Staubli VAL3: HMI_pointEdit.pjx

--- HMI_pointEdit.pjx ---
Parameters version=s8.15.3Cs9_BS3337 stackSize=5000 millimeterUnit=true
Program file=bind.pgx
Program file=insertAction.pgx
Program file=insertDelay.pgx
Program file=insertDelay1.pgx
Program file=insertIF.pgx
Program file=insertSignal.pgx
Program file=insertSwitch.pgx
Program file=load.pgx
Program file=main.pgx
Program file=onStart.pgx
Program file=paraBind.pgx
Program file=paraEdit.pgx
Program file=paraStart.pgx
Program file=refreshlist.pgx
Program file=sCommentIO.pgx
Program file=start.pgx
Program file=stop.pgx
Program file=teachPoint.pgx
Data file=HMI_pointEdit.dtx
Library alias=util path=Disk://HMI_cs9/HMI_util/HMI_util.pjx
Library alias=trajectory path=Disk://source/projectSource/trajectory/trajectory.pjx
Library alias=io path=Disk://source/projectSource/io/io.pjx
Library alias=savedata path=Disk://source/saveData/saveData.pjx
Library alias=actiondata path=Disk://data/actionData/actionData.pjx
Library alias=rs path=Disk://source/projectSource/robotStatus/robotStatus.pjx

--- HMI_pointEdit.dtx ---
mdesc mNomSpeed
bool bBack
string sTrajItem
string sUsingLib
string sUsingFrame
string sUsingTool
public bool bBool[30]
string sPageIndex
string sPageNum
public string sList = "0"
string sSelPoint
num nPageIndex
num nPageNum
bool bRefresh
bool bConfirm
bool bBackSignal
string sSignalType
string sSignalIndex
num nSignalValue
num nSignalType
string sLastType
string sIOList
bool bConfirmDelay
bool bBackDelay
num nSetDelay
public string sIFtype[3]
string sIFIndex[3]
public num nIOindex[3]
public num nIFvalue[3]
bool bConfirmIF
bool bBackIF
string sANDOR[2]
public num nANDOR[2]
num nIFtype[3]
num nParaSpeed
num nParaAccel
num nParaBlend
num nParaPercent
string sParaType
bool bParaJoint
bool bParaOFF
num nMoveType
bool bParaConfirm
bool bParaBack
bool bPAllModify
bool bLast
bool bToSave
frame fUsingFrame = {fatherId=world[0]}
tool tUsingTool = {fatherId=flange[0]}
public num nTRSF[12]
public string sTRSF[12]
string sBlendType
string sLastItem
string sLastMtype
num _nFrameID
num _nToolID
num _nPointIndex
string sComment
num nPointIndex
bool bSafePoint
string sActionList
bool bAConfirm
bool bACancel
string sSelAction
bool bConfirmSwitch
bool bBackSwitch
bool bMark
public string sCommentIO1
bool bToSave1
string sLastTrajItem
string sSelMovCPoint
bool bRecord
bool bMoveTo
bool bConfirmMovC
bool bCancelMovC
bool bShow2Point
string sParaPointType[2]

--- main.pgx ---
public program main(string x_sTrajItem)
  local bool l_bExit
  local num l_nPoint
  local bool l_bResult
  local num l_nPointSize
  local num l_nMoveType
  local bool l_bOperate
begin
  do
    if util:sPage!="point"
      util:sPage="point"
      call util:loadingPage()
      call onStart(x_sTrajItem)
      call trajectory:getFrameID(x_sTrajItem,_nFrameID)
      call trajectory:getToolID(x_sTrajItem,_nToolID)
      call refreshlist()
      call bind()
      userPage(util:sPage)
      delay(0.1)
      sLastItem=""
    endIf
    //point Move
    if workingMode()==1
      if sSelPoint!=sLastItem and sSelPoint!=""
        sLastItem=sSelPoint
        call trajectory:getPointIndex(sTrajItem,sSelPoint,l_nPoint,l_bResult)
        if !bMark
          if isPowered()
            //guohangxin modified 2023.03.23
            //            call trajectory:pointMove(sTrajItem,l_nPoint)
            if taskStatus("stepMove")>-1
              taskKill("stepMove")
              wait(taskStatus("stepMove")==-1)
            endIf
            taskCreate "stepMove",10,trajectory:pointMove(sTrajItem,l_nPoint)
          endIf
        else
          call trajectory:setMark(sTrajItem,l_nPoint)
          bRefresh=true
        endIf
      endIf
    endIf
    //button
    if bBool[0]
      //示教
      bBool[0]=false
      call trajectory:getPointIndex(sTrajItem,sSelPoint,l_nPoint,l_bResult)
      if l_bResult
        //call trajectory:teachPoint(sTrajItem,l_nPoint,bToSave)
        call teachPoint()
        bRefresh=true
      else
        userPageAlert("请选择有效点位！")
      endIf
    elseIf bBool[1]
      //标记
      bBool[1]=false
      bMark=!bMark
      if !bMark
        userPageSet("point","btn1","innerHTML","标记")
        call trajectory:resetMark(sTrajItem)
        bRefresh=true
      else
        userPageSet("point","btn1","innerHTML","取消标记")
        //call trajectory:resizeMark(sTrajItem)
      endIf
    elseIf bBool[2]
      bBool[2]=false
      //插入if
      call insertIF()
    elseIf bBool[3]
      bBool[3]=false
      //编辑
      call trajectory:getPointIndex(sTrajItem,sSelPoint,l_nPoint,l_bResult)
      if l_bResult
        call trajectory:getMoveType(sTrajItem,l_nPoint,l_nMoveType)
        if l_nMoveType==0 or l_nMoveType==1 or l_nMoveType==2
          call paraEdit()
        endIf
      else
        userPageAlert("未选择有效项！")
      endIf
    elseIf bBool[4]
      bBool[4]=false
      //插入点位
      call trajectory:getPointIndex(sTrajItem,sSelPoint,l_nPoint,l_bResult)
      if l_bResult
        call trajectory:insertPoint(sTrajItem,l_nPoint,bToSave)

      else
        call trajectory:getPointSize(sTrajItem,l_nPointSize)
        call trajectory:insertPoint(sTrajItem,l_nPointSize-1,bToSave)
      endIf
      bRefresh=true
    elseIf bBool[5]
      bBool[5]=false
      //删除
      call trajectory:getPointIndex(sTrajItem,sSelPoint,l_nPoint,l_bResult)
      if l_bResult
        call trajectory:deletePoint(sTrajItem,l_nPoint,bToSave)
      else
        userPageAlert("未选中有效点位")
      endIf
      bRefresh=true
    elseIf bBool[6]
      bBool[6]=false
      //插入信号
      call insertSignal()
      bRefresh=true
    elseIf bBool[7]
      bBool[7]=false
      //保存
      call trajectory:onSave(bToSave)
    elseIf bBool[8]
      bBool[8]=false
      //head page
      nPageIndex=0
      l_nPoint=0
      bRefresh=true
    elseIf bBool[9]
      //page up
      bBool[9]=false
      if nPageIndex>0
        nPageIndex=nPageIndex-1
        l_nPoint=0
      endIf
      bRefresh=true
    elseIf bBool[10]
      bBool[10]=false
      //page down
      if nPageIndex<nPageNum-1
        nPageIndex=nPageIndex+1
        l_nPoint=0
      endIf
      bRefresh=true
    elseIf bBool[11]
      //end page
      bBool[11]=false
      nPageIndex=nPageNum-1
      l_nPoint=0
      bRefresh=true
    elseIf bBool[12]
      bBool[12]=false
      call trajectory:getPointIndex(sTrajItem,sSelPoint,l_nPoint,l_bResult)
      if l_bResult
        call trajectory:insertENDIF(sTrajItem,l_nPoint,bToSave)
      else
        userPageAlert("未选中有效点位")
      endIf
      bRefresh=true
    elseIf bBool[13]
      bBool[13]=true
      //delay
      call insertDelay()
      bRefresh=true
    elseIf bBool[14]
      bBool[14]=false
      call trajectory:getPointIndex(sTrajItem,sSelPoint,l_nPoint,l_bResult)
      if l_bResult
        call trajectory:insertJoint(sTrajItem,l_nPoint,bToSave)
      else
        call trajectory:getPointSize(sTrajItem,l_nPointSize)
        call trajectory:insertJoint(sTrajItem,l_nPointSize-1,bToSave)
      endIf
      bRefresh=true
    elseIf bBool[15]
      bBool[15]=false
      call insertAction()
    elseIf bBool[16]
      //插入圆弧点位
      bBool[16]=false
      call trajectory:getPointIndex(sTrajItem,sSelPoint,l_nPoint,l_bResult)
      if l_bResult
        call trajectory:insertCirclePoint(sTrajItem,l_nPoint,bToSave)
      else
        userPageAlert("未选择有效项！")
      endIf
      bRefresh=true
    elseIf bBool[19]
      bBool[19]=false
      //粘贴
      call trajectory:getPointIndex(sTrajItem,sSelPoint,l_nPoint,l_bResult)
      call trajectory:copyPoint1(sTrajItem,l_nPoint)
      bMark=false
      bRefresh=true
    elseIf bBool[20]
      bBool[20]=false
      call trajectory:copyPoint(sTrajItem,bMark)
    elseIf bBool[17]
      bBool[17]=false
      call trajectory:getPointIndex(sTrajItem,sSelPoint,l_nPoint,l_bResult)
      if l_bResult
        //2025.7.21 add 喷淋delay
        call insertDelay1()
        l_nPoint=l_nPoint+1
        if l_nPoint%13==0
          nPageIndex=nPageIndex+1
        endIf
        l_bOperate=true
      else
        userPageAlert("未选中有效点位")
      endIf
      bRefresh=true
    elseIf bBack
      bBack=false

      //call trajectory:onSave(bToSave)

      l_bExit=true
    endIf

    if bRefresh
      bRefresh=false
      nPointIndex=l_nPoint
      call refreshlist()
      //      sSelPoint=sList[nPointIndex-nPageIndex*49]
      //      if sList[nPageIndex]==""
      //        sSelPoint=sList[0]
      //      endIf
    endIf
    //jogmode
    call util:jogMode(_nToolID,_nFrameID)
    //如果出现点位不可达的情况，清除当前步进任务并提示点位不可达
    //guohangxin modified 2023.03.23
    if taskStatus("stepMove")>1
      taskKill("stepMove")
      popUpMsg("当前手臂位置运动不到到步进点位")
      resetMotion()
    endIf
    delay(0)
  until l_bExit==true
  sLastTrajItem=x_sTrajItem
  if bToSave
    //bToSave=false
    l_bResult=userPageConfirm("数据已修改，是否需要保存数据？")
    if l_bResult
      call trajectory:onSave(bToSave)
    endIf
  endIf
end

--- start.pgx ---
program start()
begin
end

--- bind.pgx ---
public program bind()
  local string l_sbtn
  local num l_i
begin
  userPageBindClick("point","btnback",bBack,true)
  userPageBind("point","lbl2","innerHTML",sTrajItem,1,"r")
  userPageBind("point","lbllib","innerHTML",sUsingLib,1,"r")
  userPageBind("point","lblframe","innerHTML",sUsingFrame,1,"r")
  userPageBind("point","lbltool","innerHTML",sUsingTool,1,"r")

  userPageBind("point","lblpageindex","innerHTML",sPageIndex,1,"r")
  userPageBind("point","lblpagenum","innerHTML",sPageNum,1,"r")

  //click
  for l_i = 0 to size(bBool)-1
    l_sbtn="btn"+toString("",l_i)
    userPageBindClick("point",l_sbtn,bBool[l_i],true)
  endFor

  //lst
  //userPageBind("point","lst1","options",sList,49,"r")

  userPageBind("point","lst1","value",sSelPoint,1,"rw")
end

--- insertAction.pgx ---
public program insertAction()
  local bool l_bExit
  local num l_i
  local num l_nActionIndex
  local bool l_bResult
  local num l_nPoint
  local bool l_bResult1
begin
  do
    if util:sPage!="insertAction"
      util:sPage="insertAction"
      resize(sActionList,1,size(actiondata:aActItem))
      for l_i = 0 to size(sActionList)-1
        sActionList[l_i]=toString("",l_i)+","+actiondata:aActItem[l_i].sComment
      endFor
      sSelAction=""
      userPageBind("insertAction","cbx1","options",sActionList,size(sActionList),"r")
      userPageBind("insertAction","cbx1","value",sSelAction,1,"rw")
      userPageBindClick("insertAction","btn1",bAConfirm,true)
      userPageBindClick("insertAction","btn2",bACancel,true)
      userPage(util:sPage)
      delay(0.5)
    endIf
    //
    if bAConfirm
      bAConfirm=false
      call trajectory:getPointIndex(sTrajItem,sSelPoint,l_nPoint,l_bResult1)
      toNum(sSelAction,l_nActionIndex,l_bResult)
      if l_bResult
        call trajectory:insertAction(sTrajItem,l_nPoint,l_nActionIndex,bToSave)
        l_bExit=true
      else
        userPageAlert("选择正确的action")
      endIf
    elseIf bACancel
      bACancel=false
      l_bExit=true

    endIf

    delay(0)
  until l_bExit==true
end

--- insertDelay.pgx ---
public program insertDelay()
  local bool l_bExit
  local bool l_bResult
  local num l_nPoint
begin
  do

    if util:sPage!="insertDelay"
      util:sPage="insertDelay"
      nSetDelay=0
      userPageBindClick("insertDelay","btn1",bConfirmDelay,true)
      userPageBindClick("insertDelay","btn2",bBackDelay,true)
      userPageBind("insertDelay","nmb1","value",nSetDelay,1,"rw")
      userPage(util:sPage)
      delay(0.5)

    endIf


    if bConfirmDelay
      bConfirmDelay=false
       call trajectory:getPointIndex(sTrajItem,sSelPoint,l_nPoint,l_bResult)
      call trajectory:insertDelay(sTrajItem,l_nPoint,bToSave,7,nSetDelay)
      l_bExit=true

    elseIf bBackDelay
      bBackDelay=false
      l_bExit=true
    endIf




    delay(0)
  until l_bExit==true
end

--- insertDelay1.pgx ---
public program insertDelay1()
  local bool l_bExit
  local bool l_bResult
  local num l_nPoint
begin
  do

    //    if util:sPage!="insertDelay"
    //      util:sPage="insertDelay"
    //      nSetDelay=0
    //      userPageBindClick("insertDelay","btn1",bConfirmDelay,true)
    //      userPageBindClick("insertDelay","btn2",bBackDelay,true)
    //      userPageBind("insertDelay","nmb1","value",nSetDelay,1,"rw")
    //      userPage(util:sPage)
    //      delay(0.5)

    //    endIf

    //2024.11.20 add 插入喷淋延时由上位机控制时长s
    //    if bConfirmDelay
    //      bConfirmDelay=false
    nSetDelay=0
    call trajectory:getPointIndex(sTrajItem,sSelPoint,l_nPoint,l_bResult)
    call trajectory:insertDelay(sTrajItem,l_nPoint,bToSave,11,nSetDelay)
    l_bExit=true

    //    elseIf bBackDelay
    //      bBackDelay=false
    //      l_bExit=true
    //    endIf



    delay(0)
  until l_bExit==true
end

--- insertIF.pgx ---
program insertIF()
  local bool l_bExit
  local num l_i
  local string l_scbx
  local bool l_bResult
  local string l_snmb
  local num l_nPoint
begin
  do
    if util:sPage!="insertIF"
      util:sPage="insertIF"

      for l_i = 0 to 2
        sANDOR[0]=""
        sANDOR[1]=""
        nIOindex[l_i]=0
        nIFtype[l_i]=0
        sIFIndex[l_i]=""
        sIFtype[l_i]=""
        nIFvalue[l_i]=0
        l_scbx="cbx"+toString("",l_i)
        userPageBind("insertIF",l_scbx,"value",sIFtype[l_i],1,"rw")
        l_scbx="cbx1"+toString("",l_i)
        userPageBind("insertIF",l_scbx,"value",sIFIndex[l_i],1,"rw")
        l_snmb="nmb"+toString("",l_i)
        userPageBind("insertIF",l_snmb,"value",nIFvalue[l_i],1,"rw")
      endFor
      userPageBind("insertIF","cbx7","value",sANDOR[0],1,"rw")
      userPageBind("insertIF","cbx8","value",sANDOR[1],1,"rw")
      userPageBindClick("insertIF","btn1",bConfirmIF,true)
      userPageBindClick("insertIF","btn2",bBackIF,true)
      userPage(util:sPage)
      delay(0.5)

    endIf
    for l_i = 0 to 2
      toNum(sIFIndex[l_i],nIOindex[l_i],l_bResult)
      switch sIFtype[l_i]
        case "DIN"
          nIFtype[l_i]=1
        break
        case "DOUT"
          nIFtype[l_i]=2
        break
        case "AIN"
          nIFtype[l_i]=3
        break
        case "AOUT"
          nIFtype[l_i]=4
        break
      endSwitch
    endFor
    for l_i = 0 to 1
      switch sANDOR[l_i]
        case "AND"
          nANDOR[l_i]=1
        break
        case "OR"
          nANDOR[l_i]=2
        break
        default
          nANDOR[l_i]=0
        break
      endSwitch
    endFor
    //button
    if bConfirmIF
      bConfirmIF=false
       call trajectory:getPointIndex(sTrajItem,sSelPoint,l_nPoint,l_bResult)

      call trajectory:insertIF(sTrajItem,l_nPoint,nIFtype,nIOindex,nIFvalue,nANDOR,bToSave)
      l_bExit=true
    elseIf bBackIF
      bBackIF=false
      l_bExit=true
    endIf






    delay(0)
  until l_bExit==true
end

--- insertSignal.pgx ---
public program insertSignal()
  local bool l_bExit
  local bool l_bResult
  local num l_nPoint
  local bool l_bResult1
  local num l_nIndex
begin
  do
    if util:sPage!="insertSignal"
      util:sPage="insertSignal"
      sSignalType=""
      sSignalIndex=""
      nSignalValue=0

      userPageBindClick("insertSignal","btn1",bConfirm,true)
      userPageBindClick("insertSignal","btn2",bBackSignal,true)
      userPageBind("insertSignal","cbx1","value",sSignalType,1,"rw")
      userPageBind("insertSignal","cbx2","value",sSignalIndex,1,"rw")
      userPageBind("insertSignal","nmb1","value",nSignalValue,1,"rw")

      userPage(util:sPage)
      delay(0.5)
      sLastType=""
    endIf
    //
    if sSignalType!=sLastType
      sLastType=sSignalType
      switch sSignalType
        case "DIN","DOUT"
          resize(sIOList,1,1)
          sIOList=""
          //userPageUnbind("insertSignal","cbx2","options")
        break
        case "AIN"
          call io:setAngINList(sIOList)
          // userPageBind("insertSignal","cbx2","options",sIOList,size(sIOList),"r")
        break
        case "AOUT"
          call io:setAngOUTList(sIOList)
          //userPageBind("insertSignal","cbx2","options",sIOList,size(sIOList),"r")
        break
      endSwitch
      switch sSignalType
        case "DIN"
          nSignalType=3
        break
        case "DOUT"
          nSignalType=4
        break
        case "AIN"
          nSignalType=5
        break
        case "AOUT"
          nSignalType=6
        break
        default
          nSignalType=0
        break
      endSwitch


    endIf
    //signal type



    //btn
    if bConfirm
      bConfirm=false
      call trajectory:getPointIndex(sTrajItem,sSelPoint,l_nPoint,l_bResult)
      toNum(sSignalIndex,l_nIndex,l_bResult1)
      if l_nIndex>io:nMaxAnalog-1 and (nSignalType==5 or nSignalType==6)
        userPageAlert("信号索引大于模拟量最大个数")
      else
        call trajectory:insertSignal(sTrajItem,l_nPoint,bToSave,nSignalType,l_nIndex,nSignalValue)
        l_bExit=true
      endIf


    elseIf bBackSignal
      bBackSignal=false
      l_bExit=true
    endIf

    //

    delay(0)
  until l_bExit==true
end

--- insertSwitch.pgx ---
public program insertSwitch()
begin
  //   do

  //    if util:sPage!="insertSwitch"
  //      util:sPage="insertSwitch"

  //      userPageBindClick("insertDelay","btn1",bConfirmSwitch,true)
  //      userPageBindClick("insertDelay","btn2",bBackSwitch,true)
  //      userPageBind("insertSwitch","cbx2","options",nSetDelay,1,"rw")
  //      userPage(util:sPage)
  //      delay(0.5)

  //    endIf


  //    if bConfirmDelay
  //      bConfirmDelay=false
  //       call trajectory:getPointIndex(sTrajItem,sSelPoint,l_nPoint,l_bResult)
  //      call trajectory:insertDelay(sTrajItem,l_nPoint,bToSave,7,nSetDelay)
  //      l_bExit=true

  //    elseIf bBackDelay
  //      bBackDelay=false
  //      l_bExit=true
  //    endIf




  //    delay(0)
  //  until l_bExit==true
end

--- load.pgx ---
program load()
  local string l_sPath
  local bool l_bResult
  local num l_nResult
begin
//call trajectory:loadTRAJ(savedata:nLibIndex,l_nResult)
end

--- onStart.pgx ---
public program onStart(string x_sTrajItem)
  local num l_i
  local num l_nFrameID
  local num l_nToolID
  local num l_nLibNum
  local bool l_bResult
begin
  if sLastTrajItem!=x_sTrajItem
    nPageIndex=0
    nPointIndex=0
  endIf
  call load()
  //
  delay(0)
  sTrajItem=x_sTrajItem
  //

  bBack=false
  for l_i = 0 to size(bBool)-1
    bBool[l_i]=false
  endFor
  //
  for l_i = 0 to size(sList)-1
    sList[l_i]=""
  endFor
  //
  call trajectory:getFrameID(sTrajItem,l_nFrameID)
  call trajectory:getToolID(sTrajItem,l_nToolID)
  call trajectory:getLibName(l_nLibNum,l_bResult)
  call savedata:getFrame(l_nFrameID,fUsingFrame)
  call savedata:getTool(l_nToolID,tUsingTool)
  $jogContext(tUsingTool,fUsingFrame,0)

  sUsingFrame=toString("",l_nFrameID)
  sUsingTool=toString("",l_nToolID)
  sUsingLib=toString("",l_nLibNum)
  logMsg("<traj-jogContext> tool:"+sUsingTool+",frame:"+sUsingFrame)

  sSelPoint=""
  bMark=false



end

--- paraBind.pgx ---
public program paraBind()
  local num l_i
  local string l_snmb
  local string l_slbl
begin
  //  userPageBind("paraEdit","nmb1","value",nParaSpeed,1,"rw")
  //  userPageBind("paraEdit","nmb2","value",nParaAccel,1,"rw")
  //  userPageBind("paraEdit","nmb3","value",nParaBlend,1,"rw")
  //  userPageBind("paraEdit","nmb4","value",nParaPercent,1,"rw")
  //  for l_i = 0 to 5
  //    l_snmb="nmb5"+toString("",l_i)
  //    userPageBind("paraEdit",l_snmb,"value",nTRSF[l_i],1,"rw")
  //    l_slbl="lbl5"+toString("",l_i)
  //    userPageBind("paraEdit",l_slbl,"innerHTML",sTRSF[l_i],1,"r")
  //  endFor
  //  //cbx
  //  userPageBind("paraEdit","cbx1","value",sParaType,1,"rw")
  //  //chk
  //  userPageBind("paraEdit","cbx3","value",sBlendType,1,"rw")
  //  //button
  //  userPageBindClick("paraEdit","btn1",bParaConfirm,true)
  //  userPageBindClick("paraEdit","btn2",bParaBack,true)
  //  userPageBindClick("paraEdit","btn3",bPAllModify,true)
  //  //txt1
  //  userPageBind("paraEdit","txt1","value",sComment,1,"rw")

  //  //chk
  //  userPageBind("paraEdit","chk1","checked",bSafePoint,1,"rw")

  userPageBind("paraEdit","nmb1","value",nParaSpeed,1,"rw")
  userPageBind("paraEdit","nmb2","value",nParaAccel,1,"rw")
  userPageBind("paraEdit","nmb3","value",nParaBlend,1,"rw")
  userPageBind("paraEdit","nmb4","value",nParaPercent,1,"rw")
  for l_i = 0 to 9
    l_snmb="nmb5"+toString("",l_i)
    userPageBind("paraEdit",l_snmb,"value",nTRSF[l_i],1,"rw")
    l_slbl="lbl5"+toString("",l_i)
    userPageBind("paraEdit",l_slbl,"innerHTML",sTRSF[l_i],1,"r")
  endFor
  for l_i = 0 to 1
    l_snmb="nmb6"+toString("",l_i)
    userPageBind("paraEdit",l_snmb,"value",nTRSF[l_i+10],1,"rw")
    l_slbl="lbl6"+toString("",l_i)
    userPageBind("paraEdit",l_slbl,"innerHTML",sTRSF[l_i+10],1,"r")
  endFor
  //cbx
  userPageBind("paraEdit","cbx1","options",sParaPointType,size(sParaPointType),"r")
  userPageBind("paraEdit","cbx1","value",sParaType,1,"rw")
  //chk
  userPageBind("paraEdit","cbx3","value",sBlendType,1,"rw")
  //button
  userPageBindClick("paraEdit","btn1",bParaConfirm,true)
  userPageBindClick("paraEdit","btn2",bParaBack,true)
  userPageBindClick("paraEdit","btn3",bPAllModify,true)
  //txt1
  userPageBind("paraEdit","txt1","value",sComment,1,"rw")

  //chk
  userPageBind("paraEdit","chk1","checked",bSafePoint,1,"rw")
end

--- paraEdit.pgx ---
public program paraEdit()
  local num l_nPoint
  local bool l_bResult
  local bool l_bExit
  local num l_i
  local string l_snmb
  local string l_slbl
begin
  call trajectory:getPointIndex(sTrajItem,sSelPoint,_nPointIndex,l_bResult)
  if l_bResult

    do
      if util:sPage!="paraEdit"
        util:sPage="paraEdit"
        call paraStart(_nPointIndex)
        call paraBind()
        userPage(util:sPage)
        delay(0.5)
        //sLastMtype=""
        sLastType=""
      endIf

      if sParaType!=sLastType and sParaType!=""
        sLastType=sParaType
        call trajectory:pointEditValue(sParaType,sTrajItem,_nPointIndex,nTRSF,sTRSF,bShow2Point)
        call paraBind()
      endIf

      if sParaType=="POINT" or sParaType==""
        nMoveType=1
      elseIf sParaType=="JOINT"
        nMoveType=0
      elseIf sParaType=="CIRCLE"
        nMoveType=2
      endIf

      //button
      if bParaConfirm
        bParaConfirm=false
        //call trajectory:getPointIndex(sTrajItem,sSelPoint,_nPointIndex,l_bResult)
        call trajectory:modifyPara(sTrajItem,_nPointIndex,nMoveType,nParaSpeed,nParaBlend,nParaPercent,sComment,bSafePoint,sBlendType,bToSave,nTRSF,nParaAccel)

        l_bExit=true
      elseIf bPAllModify
        bPAllModify=false
        //call trajectory:getPointIndex(sTrajItem,sSelPoint,_nPointIndex,l_bResult)
        call trajectory:modifyAll(sTrajItem,nMoveType,nParaSpeed,nParaBlend,nParaPercent,sBlendType,bToSave,nParaAccel)
        l_bExit=true
      elseIf bParaBack
        bParaBack=false
        l_bExit=true
      endIf
      delay(0)
    until l_bExit==true
    //    l_bResult=userPageConfirm("数据已修改，是否需要保存数据？")
    //    if l_bResult
    //      call trajectory:onSave(bToSave)
    //    endIf
  else
    userPageAlert("未选择有效点位！")
  endIf
end

--- paraStart.pgx ---
program paraStart(num x_nPoint)
begin

  //  call trajectory:getPointPara(sTrajItem,x_nPoint,nMoveType,nParaSpeed,nParaAccel,nParaBlend,nParaPercent,sComment,bSafePoint,sBlendType,nTRSF,sTRSF)
  //  switch nMoveType
  //    case 0
  //      sParaType="POINT"
  //    break
  //    case 1
  //      sParaType="JOINT"
  //    break
  //  endSwitch

  call trajectory:getPointPara(sTrajItem,x_nPoint,nMoveType,nParaSpeed,nParaAccel,nParaBlend,nParaPercent,sComment,bSafePoint,sBlendType,nTRSF,sTRSF)
  switch nMoveType
    case 1
      bShow2Point=false
      resize(sParaPointType,1,2)
      sParaPointType[0]="POINT"
      sParaPointType[1]="JOINT"
      sParaType="POINT"
    break
    case 0
      bShow2Point=false
      resize(sParaPointType,1,2)
      sParaPointType[0]="POINT"
      sParaPointType[1]="JOINT"
      sParaType="JOINT"
    break
    case 2
      bShow2Point=true
      resize(sParaPointType,1,1)
      sParaPointType[0]="CIRCLE"
      sParaType="CIRCLE"
    break
  endSwitch
end

--- refreshlist.pgx ---
public program refreshlist()
  local num l_nSize
  local string l_sMsg
  local num l_i
  local num l_nPointSize
  local num l_nPoint
  local bool l_bResult
begin
  call trajectory:getPointSize(sTrajItem,l_nPointSize)

  //page
  if l_nPointSize<50
    nPageNum=1
  else
    nPageNum=roundUp(l_nPointSize/49)
  endIf

  if nPageNum==1
    resize(sList,1,l_nPointSize)
    for l_i = 0 to size(sList)-1
      call trajectory:pointToString(l_sMsg,sTrajItem,l_i+49*nPageIndex)
      sList[l_i]=toString("",l_i+49*nPageIndex)+l_sMsg
    endFor
  else
    if nPageIndex<nPageNum-1
      resize(sList,1,49)
      for l_i = 0 to 48
        call trajectory:pointToString(l_sMsg,sTrajItem,l_i+49*nPageIndex)
        sList[l_i]=toString("",l_i+49*nPageIndex)+l_sMsg
      endFor
    else
      if l_nPointSize%49==0
        resize(sList,1,49)
      else
        resize(sList,1,l_nPointSize%49)
      endIf
      for l_i = 0 to size(sList)-1
        call trajectory:pointToString(l_sMsg,sTrajItem,l_i+49*nPageIndex)
        sList[l_i]=toString("",l_i+49*nPageIndex)+l_sMsg
      endFor

    endIf
  endIf
  userPageBind("point","lst1","options",sList,size(sList),"r")
  sPageIndex=toString("",nPageIndex+1)
  sPageNum=toString("",nPageNum)
  //
  //  if nPageIndex>(nPageNum-1)
  //    nPageIndex=(nPageNum-1)
  //  endIf
  //  //slist
  //  if nPageIndex==(nPageNum-1)
  //    if l_nPointSize%49==0
  //      l_nSize=49
  //    else
  //      l_nSize=l_nPointSize%49
  //    endIf
  //    for l_i = 0 to l_nSize-1
  //      call trajectory:pointToString(l_sMsg,sTrajItem,l_i+49*nPageIndex)
  //      sList[l_i]=toString("",l_i+49*nPageIndex)+l_sMsg
  //    endFor
  //    if l_nSize<49
  //      for l_i= l_nSize to 48
  //        sList[l_i]=""
  //      endFor
  //    endIf
  //  else
  //    for l_i = 0 to size(sList)-1
  //      call trajectory:pointToString(l_sMsg,sTrajItem,l_i+49*nPageIndex)
  //      sList[l_i]=toString("",l_i+49*nPageIndex)+l_sMsg
  //    endFor
  //  endIf
  //  sPageIndex=toString("",nPageIndex+1)
  //  sPageNum=toString("",nPageNum)
  //  //sSelPoint=sList[nPointIndex-nPageIndex*49]
end

--- sCommentIO.pgx ---
program sCommentIO()
begin
end

--- stop.pgx ---
program stop()
begin
end

--- teachPoint.pgx ---
program teachPoint()
  local num l_nPoint
  local bool l_bResult
  local num l_nMoveType
  local bool l_bExit
begin
  //2024.12.23 add 增加movec示教界面
  call trajectory:getPointIndex(sTrajItem,sSelPoint,l_nPoint,l_bResult)
  call trajectory:getMoveType(sTrajItem,l_nPoint,l_nMoveType)
  call trajectory:getFrameID(sTrajItem,_nFrameID)
  call trajectory:getToolID(sTrajItem,_nToolID)
  if l_bResult
    if l_nMoveType==0 or l_nMoveType==1
      //moveL、moveJ示教
      call trajectory:teachPoint(sTrajItem,l_nPoint,bToSave)
    elseIf l_nMoveType==2
      //进入moveC示教界面
      do
        if util:sPage!="movecTeach"
          util:sPage="movecTeach"
          sSelMovCPoint="中间点"
          userPageBindClick("movecTeach","btn1",bRecord,true)
          userPageBindClick("movecTeach","btn2",bMoveTo,true)
          userPageBindClick("movecTeach","btn3",bConfirmMovC,true)
          userPageBindClick("movecTeach","btn4",bCancelMovC,true)
          userPage(util:sPage)
          delay(0.2)
        endIf

        if bRecord
          bRecord=false
          if sSelMovCPoint=="中间点"
            call trajectory:teachPoint1(sTrajItem,l_nPoint,0)
            popUpMsg("圆弧中间点记录完成！")
          elseIf sSelMovCPoint=="结束点"
            call trajectory:teachPoint1(sTrajItem,l_nPoint,1)
            popUpMsg("圆弧结束点记录完成！")
          endIf
        elseIf bMoveTo
          bMoveTo=false
          if sSelMovCPoint=="中间点"
            call trajectory:pointMove1(sTrajItem,l_nPoint,0)
          elseIf sSelMovCPoint=="结束点"
            call trajectory:pointMove1(sTrajItem,l_nPoint,1)
          endIf
        elseIf bConfirmMovC
          bConfirmMovC=false
          bToSave=true
          l_bExit=true
        elseIf bCancelMovC
          bCancelMovC=false
          l_bExit=true
        endIf

        //jogmode
        call util:jogMode(_nToolID,_nFrameID)
        delay(0)
      until l_bExit==true
    endIf
  else
    userPageAlert("未选择有效点位！")
  endIf
end
